(* IEC 61131-3 sources: plc-vscode/tests/st/all/rusty/tests/lit/single/stdlib_overflow, 14 files *)

(* ---- sub32_ffi_return_byte.st ---- *)
// RUN: (%COMPILE %s && %RUN) | %CHECK %s
// Stress test for u8 (BYTE) FFI return values. ROL__BYTE / ROR__BYTE in the
// Rust stdlib take and return u8. Under the target-aware extension gate
// (#1146 follow-up), the rusty side either emits `zeroext i8` on both call
// and declaration (x86 family / Darwin) or skips the attribute entirely
// (AAPCS aarch64-linux). Either way the runtime behaviour must match the
// IEC semantics: BYTE 0xFF rotated by 0 stays 0xFF; rotating 0x80 left by
// one wraps to 0x01.

FUNCTION main : DINT
VAR
    r1 : BYTE;
    r2 : BYTE;
    r3 : BYTE;
    r4 : BYTE;
END_VAR
    r1 := ROL(BYTE#16#FF, 0);
    // CHECK: 255
    printf('%d$N', r1);

    r2 := ROL(BYTE#16#80, 1);
    // CHECK: 1
    printf('%d$N', r2);

    r3 := ROR(BYTE#16#01, 1);
    // CHECK: 128
    printf('%d$N', r3);

    r4 := ROR(BYTE#16#FF, 4);
    // CHECK: 255
    printf('%d$N', r4);

    main := 0;
END_FUNCTION

(* ---- sub32_ffi_return_signed.st ---- *)
// RUN: (%COMPILE %s && %RUN) | %CHECK %s
// Stress test for the sub-32-bit FFI integer ABI fix (#1146).
// Calls Rust stdlib `MUL_LTIME` with negative `SINT` arguments and asserts
// the i8 sign-extension on the parameter side reaches the callee correctly
// under release optimizations. The original repro: passing SINT#-120 used
// to read with the upper bits unset on x86_64 release; this test pins the
// fix and lets the matching CI lanes prove the target-aware gate is right.

FUNCTION main : DINT
VAR
    a : LTIME;
    b : LTIME;
    c : LTIME;
END_VAR
    a := MUL_LTIME(LTIME#1d, SINT#-120);
    // CHECK: -10368000000000000
    printf('%lld$N', a);

    b := MUL_LTIME(LTIME#1d, SINT#-1);
    // CHECK: -86400000000000
    printf('%lld$N', b);

    c := MUL_LTIME(LTIME#1d, SINT#127);
    // CHECK: 10972800000000000
    printf('%lld$N', c);

    main := 0;
END_FUNCTION

(* ---- sub32_ffi_return_word.st ---- *)
// RUN: (%COMPILE %s && %RUN) | %CHECK %s
// Stress test for u16 (WORD) FFI return values. Same shape as the BYTE
// regression but at i16 width — exercises the second sub-32-bit slot the
// extension gate must handle consistently across targets.

FUNCTION main : DINT
VAR
    r1 : WORD;
    r2 : WORD;
    r3 : WORD;
END_VAR
    r1 := ROL(WORD#16#FFFF, 0);
    // CHECK: 65535
    printf('%d$N', r1);

    r2 := ROL(WORD#16#8000, 1);
    // CHECK: 1
    printf('%d$N', r2);

    r3 := ROR(WORD#16#0001, 1);
    // CHECK: 32768
    printf('%d$N', r3);

    main := 0;
END_FUNCTION

(* ---- add_time_overflow.st ---- *)
// RUN: (%COMPILE %s && %RUN) | %CHECK %s
// XFAIL: *
// Test that ADD with TIME overflow causes a panic

PROGRAM main
VAR
    a : TIME;
END_VAR
    // Adding 1ms to max TIME value should overflow and panic
    a := ADD(TIME#9223372036854775807ms, TIME#1ms);
    // CHECK: Should not reach here
    printf('Should not reach here$N');
END_PROGRAM

(* ---- div_time_by_lreal_zero.st ---- *)
// RUN: (%COMPILE %s && %RUN) | %CHECK %s
// XFAIL: *
// Test that DIV with TIME by LREAL zero causes a panic

PROGRAM main
VAR
    a : TIME;
END_VAR
    // Dividing TIME by zero (LREAL) should panic
    a := DIV(TIME#10ns, LREAL#0.0);
    // CHECK: Should not reach here
    printf('Should not reach here$N');
END_PROGRAM

(* ---- div_time_by_real_zero.st ---- *)
// RUN: (%COMPILE %s && %RUN) | %CHECK %s
// XFAIL: *
// Test that DIV with TIME by REAL zero causes a panic

PROGRAM main
VAR
    a : TIME;
END_VAR
    // Dividing TIME by zero (REAL) should panic
    a := DIV(TIME#10ns, REAL#0.0);
    // CHECK: Should not reach here
    printf('Should not reach here$N');
END_PROGRAM

(* ---- div_time_by_zero.st ---- *)
// RUN: (%COMPILE %s && %RUN) | %CHECK %s
// XFAIL: *
// Test that DIV with TIME by zero causes a panic

PROGRAM main
VAR
    a : TIME;
END_VAR
    // Dividing TIME by zero should panic
    a := DIV(TIME#10ns, LINT#0);
    // CHECK: Should not reach here
    printf('Should not reach here$N');
END_PROGRAM

(* ---- mul_time_lreal_overflow.st ---- *)
// RUN: (%COMPILE %s && %RUN) | %CHECK %s
// XFAIL: *
// Test that MUL with TIME and LREAL overflow causes a panic

PROGRAM main
VAR
    a : TIME;
END_VAR
    // Multiplying TIME by large LREAL value should overflow and panic
    a := MUL(TIME#-2s700ms, LREAL#3.40282347e38);
    // CHECK: Should not reach here
    printf('Should not reach here$N');
END_PROGRAM

(* ---- mul_time_real_overflow.st ---- *)
// RUN: (%COMPILE %s && %RUN) | %CHECK %s
// XFAIL: *
// Test that MUL with TIME and REAL overflow causes a panic

PROGRAM main
VAR
    a : TIME;
END_VAR
    // Multiplying TIME by max REAL value should overflow and panic
    a := MUL(TIME#-2s700ms, REAL#3.40282347e38);
    // CHECK: Should not reach here
    printf('Should not reach here$N');
END_PROGRAM

(* ---- mul_time_signed_overflow.st ---- *)
// RUN: (%COMPILE %s && %RUN) | %CHECK %s
// XFAIL: *
// Test that MUL with TIME and signed integer overflow causes a panic

PROGRAM main
VAR
    a : TIME;
END_VAR
    // Multiplying TIME by max LINT value should overflow and panic
    a := MUL(TIME#10ns, LINT#9223372036854775807);
    // CHECK: Should not reach here
    printf('Should not reach here$N');
END_PROGRAM

(* ---- mul_time_unsigned_overflow.st ---- *)
// RUN: (%COMPILE %s && %RUN) | %CHECK %s
// XFAIL: *
// Test that MUL with TIME and unsigned integer overflow causes a panic

PROGRAM main
VAR
    a : TIME;
END_VAR
    // Multiplying TIME by max ULINT value should overflow and panic
    a := MUL(TIME#1ns, ULINT#9223372036854775808);
    // CHECK: Should not reach here
    printf('Should not reach here$N');
END_PROGRAM

(* ---- right_string_substring_too_long.st ---- *)
// RUN: (%COMPILE %s && %RUN 2>&1) | %CHECK %s
// XFAIL: *
// Test that RIGHT with substring length > string length causes a panic
// Expected failure message: Requested substring length exceeds string length.
// CHECK: Requested substring length exceeds string length.

PROGRAM main
VAR
    s : STRING;
END_VAR
    s := 'sample text';
    // Length 12 exceeds string length 11 -> should panic
    s := RIGHT(s, 12);
    // CHECK: Should not reach here
    printf('Should not reach here$N');
END_PROGRAM

(* ---- right_wstring_substring_too_long.st ---- *)
// RUN: (%COMPILE %s && %RUN 2>&1) | %CHECK %s
// XFAIL: *
// Test that RIGHT with substring length > string length causes a panic
// Expected failure message: Requested substring length exceeds string length.
// CHECK: Requested substring length exceeds string length.

PROGRAM main
VAR
    s : WSTRING;
END_VAR
    s := "sa𝄞ple text";
    // Length 12 exceeds string length 11 -> should panic
    s := RIGHT(s, 12);
    // CHECK: Should not reach here
    printf('Should not reach here$N');
END_PROGRAM

(* ---- sub_time_overflow.st ---- *)
// RUN: (%COMPILE %s && %RUN) | %CHECK %s
// XFAIL: *
// Test that SUB with TIME overflow causes a panic

PROGRAM main
VAR
    a : TIME;
END_VAR
    // Subtracting from minimum TIME value should overflow and panic
    a := SUB(TIME#-9223372036854775807ms, TIME#1ms);
    // CHECK: Should not reach here
    printf('Should not reach here$N');
END_PROGRAM
